// SIMATIC S7-200 project (STEP 7-Micro/WIN), CPU 224XP CN REL 02.01

SYMBOL_TABLE USER1
Pos_Real         VD100    // Posicion real en cuentas de encoder (REAL)
Setpoint         VD112    // Posicion objetivo de referencia en cuentas (REAL)
Accion_Control   VD116    // Accion de control calculada u (REAL)
K1               VD120    // Ganancia de posicion del controlador (97.7436) (REAL)
K2               VD124    // Ganancia de velocidad del controlador (25.8460) (REAL)
U_Abs            VD128    // Magnitud absoluta de la accion de control (REAL)
N                VD132    // Ganancia de precompensacion de la referencia (REAL)
Setpoint_In      VD136    // Referencia dinamica de posicion desde HMI (REAL)
Pos_Est          VD140    // Posicion estimada por el observador (REAL)
Vel_Est          VD144    // Velocidad estimada por el observador (REAL)
Error_Est        VD148    // Error de estimacion de la posicion ey (REAL)
L1               VD152    // Ganancia de observador para canal de posicion (0.1919) (REAL)
L2               VD156    // Ganancia de observador para canal de velocidad (0.6113) (REAL)
Phi12            VD160    // Matriz de transicion de estado elemento 12 (0.009814) (REAL)
Phi22            VD164    // Matriz de transicion de estado elemento 22 (0.963062) (REAL)
Gamma1           VD168    // Matriz de entrada elemento 1 (0.000008) (REAL)
Gamma2           VD172    // Matriz de entrada elemento 2 (0.001611) (REAL)
Pos_Est_Next     VD176    // Valor intermedio de posicion estimada siguiente (REAL)
Vel_Est_Next     VD180    // Valor intermedio de velocidad estimada siguiente (REAL)
Seta_Emergencia  I1.4     // Entrada de seguridad NC (1=OK
Variador_Run     Q0.0     // Mando Marcha/Paro del variador (1=Run
Variador_Dir     Q0.1     // Mando Direccion del variador (0=FWD
Salida_Analog    AQW0     // Consigna analoga de velocidad para el variador (0-32000)
Log_Pointer      VD400    // Puntero de escritura en la memoria de registro (DWORD)
Log_SampleCount  VW404    // Contador de muestras registradas de 0 a 200 (INT)
Log_DecimCount   VW406    // Contador de decimacion para muestreo de 50ms (INT)
Log_Active       V408.0   // Bandera de registro activo en ejecucion (BOOL)
Log_Trigger      V408.1   // Gatillo de inicio de registro manual (BOOL)
END_SYMBOL_TABLE

SYMBOL_TABLE S7-200 Symbols
Always_On        SM0.0    // 始终接通为 ON
First_Scan_On    SM0.1    // 仅第一个扫描周期中接通为 ON
Time_0_Intrvl    SMB34    // 定时中断 0 的时间间隔（从 1 至 255，以 1 毫秒为增量）。
HSC0_Ctrl        SMB37    // HSC0 设置与控制
HSC0_CV          SMD38    // HSC0 的新当前值
HSC0_PV          SMD42    // HSC0 的新预置值
END_SYMBOL_TABLE

ORGANIZATION_BLOCK MAIN:OB1
TITLE=
BEGIN
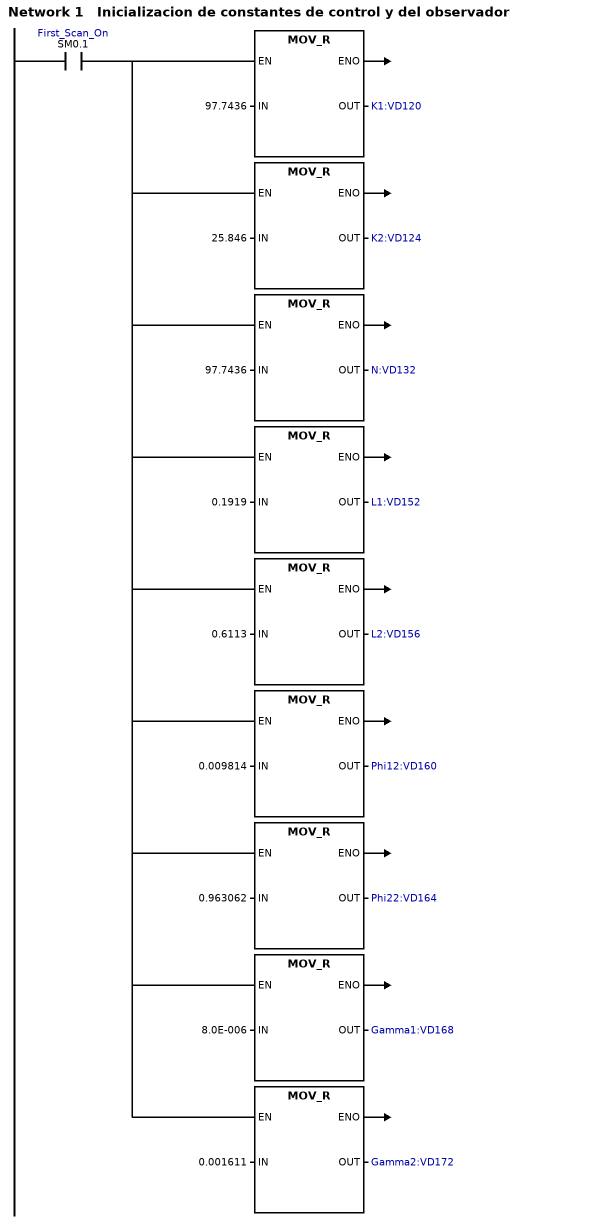
Network 1 //  Inicializacion de constantes de control y del observador
// K1
// K2
// N (Pre-compensacion)
// L1 (Ganancia de observador 1)
// L2 (Ganancia de observador 2)
// Phi12
// Phi22
// Gamma1
// Gamma2
LD     First_Scan_On:SM0.1
MOVR   97.7436, K1:VD120
MOVR   25.846, K2:VD124
MOVR   97.7436, N:VD132
MOVR   0.1919, L1:VD152
MOVR   0.6113, L2:VD156
MOVR   0.009814, Phi12:VD160
MOVR   0.963062, Phi22:VD164
MOVR   8.0E-006, Gamma1:VD168
MOVR   0.001611, Gamma2:VD172
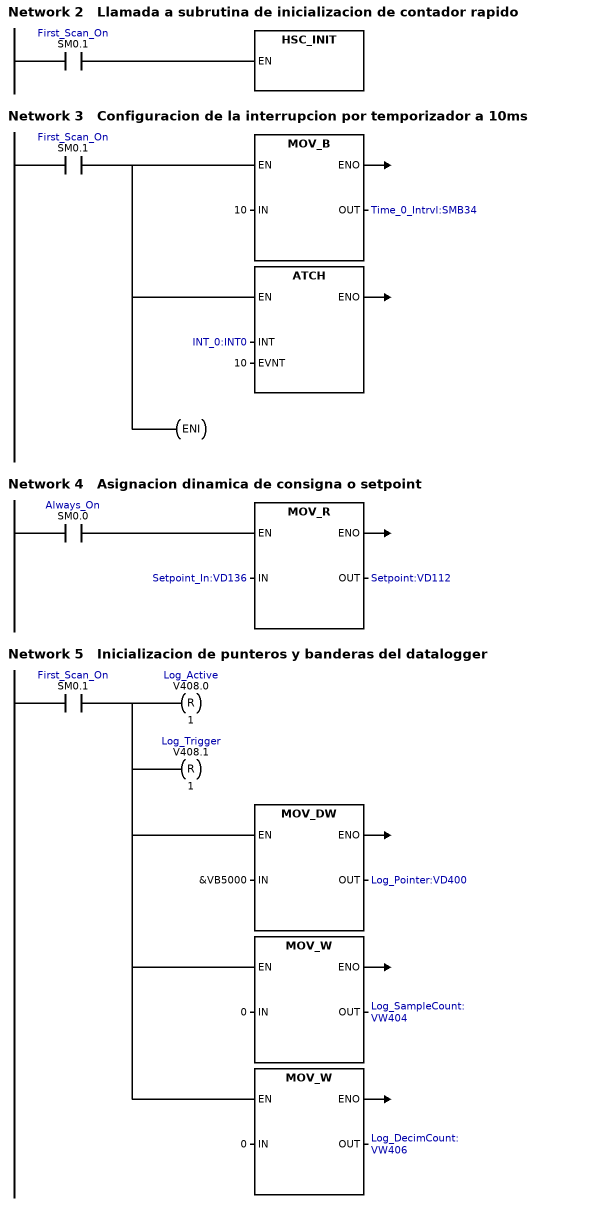
Network 2 //  Llamada a subrutina de inicializacion de contador rapido
// Llamada a SBR1 (HSC_INIT)
LD     First_Scan_On:SM0.1
CALL   HSC_INIT:SBR1
Network 3 //  Configuracion de la interrupcion por temporizador a 10ms
// Intervalo de interrupcion de 10ms
// Asociar INT0 al evento de temporizador 0
// Habilitar interrupciones globalmente
LD     First_Scan_On:SM0.1
MOVB   10, Time_0_Intrvl:SMB34
ATCH   INT_0:INT0, 10
ENI
Network 4 //  Asignacion dinamica de consigna o setpoint
// VD112 = Setpoint (Referencia)
LD     Always_On:SM0.0
MOVR   Setpoint_In:VD136, Setpoint:VD112
Network 5 //  Inicializacion de punteros y banderas del datalogger
// Desactivar bandera de datalogger activo
// Desactivar bandera de disparo (trigger)
// Direccion inicial del bufer en puntero
// Resetear contador de muestras
// Resetear contador de decimacion
LD     First_Scan_On:SM0.1
R      Log_Active:V408.0, 1
R      Log_Trigger:V408.1, 1
MOVD   &VB5000, Log_Pointer:VD400
MOVW   0, Log_SampleCount:VW404
MOVW   0, Log_DecimCount:VW406
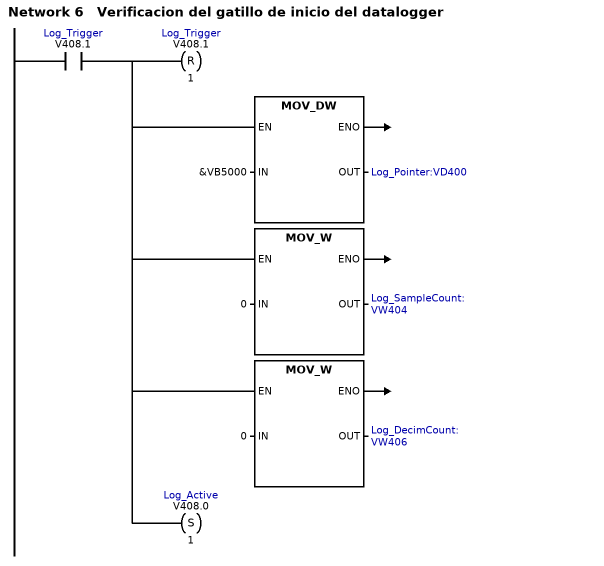
Network 6 //  Verificacion del gatillo de inicio del datalogger
// Si el usuario activa el gatillo
// Resetear bandera de gatillo
// Apuntar puntero al inicio VB5000
// Resetear contador de muestras
// Resetear contador de decimacion
// Activar bandera de datalogger activo
LD     Log_Trigger:V408.1
R      Log_Trigger:V408.1, 1
MOVD   &VB5000, Log_Pointer:VD400
MOVW   0, Log_SampleCount:VW404
MOVW   0, Log_DecimCount:VW406
S      Log_Active:V408.0, 1
END_ORGANIZATION_BLOCK

SUBROUTINE_BLOCK SBR_0:SBR0
TITLE=
BEGIN
Network 1
LD     Always_On:SM0.0
END_SUBROUTINE_BLOCK

SUBROUTINE_BLOCK HSC_INIT:SBR1
TITLE=
BEGIN
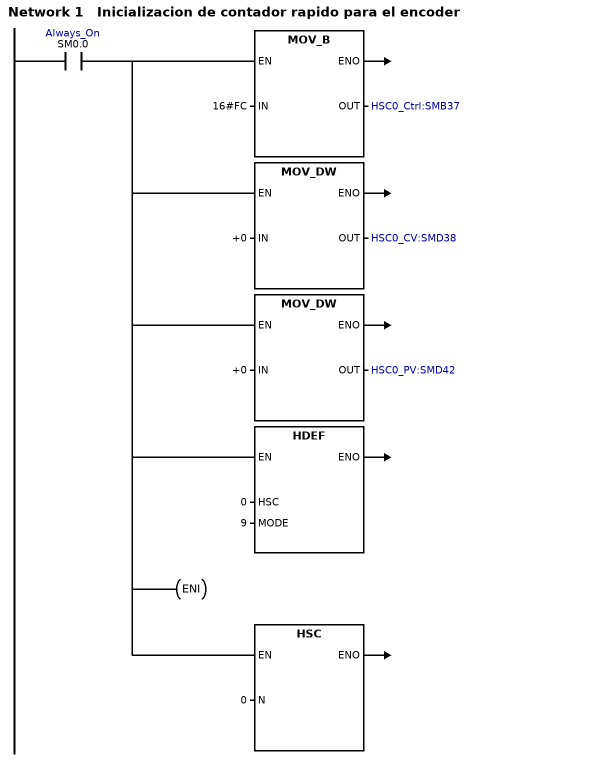
Network 1 //  Inicializacion de contador rapido para el encoder
// Configuracion de conteo: UP, 1X, habilitado
// Cargar valor actual (CV = 0)
// Cargar valor de preseleccion (PV = 0)
// Configurar HSC0 en Modo 9 (Fases A/B)
// Habilitar interrupciones
// Iniciar contador rapido HSC0
LD     Always_On:SM0.0
MOVB   16#FC, HSC0_Ctrl:SMB37
MOVD   +0, HSC0_CV:SMD38
MOVD   +0, HSC0_PV:SMD42
HDEF   0, 9
ENI
HSC    0
END_SUBROUTINE_BLOCK

INTERRUPT_BLOCK INT_0:INT0
TITLE=
BEGIN
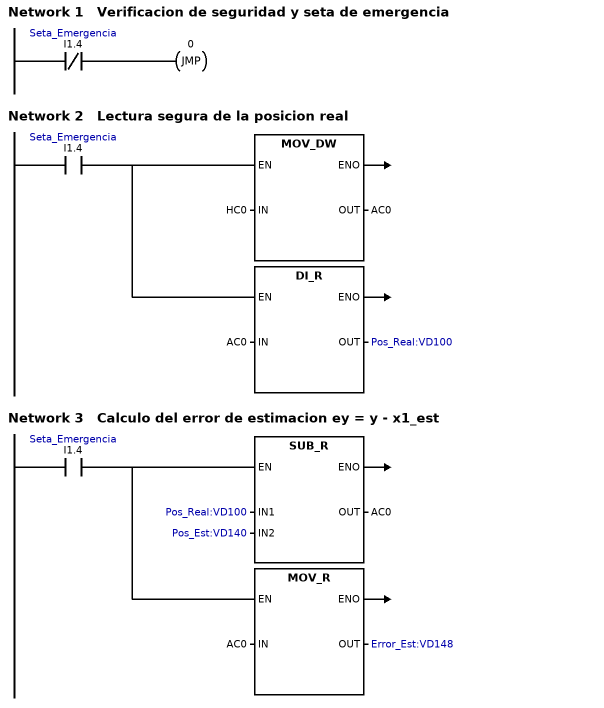
Network 1 //  Verificacion de seguridad y seta de emergencia
// Si la seta de emergencia se activa (NC abierto)
// Saltar a la etiqueta de parada segura
LDN    Seta_Emergencia:I1.4
JMP    0
Network 2 //  Lectura segura de la posicion real
// Mover lectura de HC0 a AC0
// Convertir entero de AC0 a REAL en VD100 (y)
LD     Seta_Emergencia:I1.4
MOVD   HC0, AC0
DTR    AC0, Pos_Real:VD100
Network 3 //  Calculo del error de estimacion ey = y - x1_est
// AC0 = y
// AC0 = y - x1_est
// VD148 = ey
LD     Seta_Emergencia:I1.4
MOVR   Pos_Real:VD100, AC0
-R     Pos_Est:VD140, AC0
MOVR   AC0, Error_Est:VD148
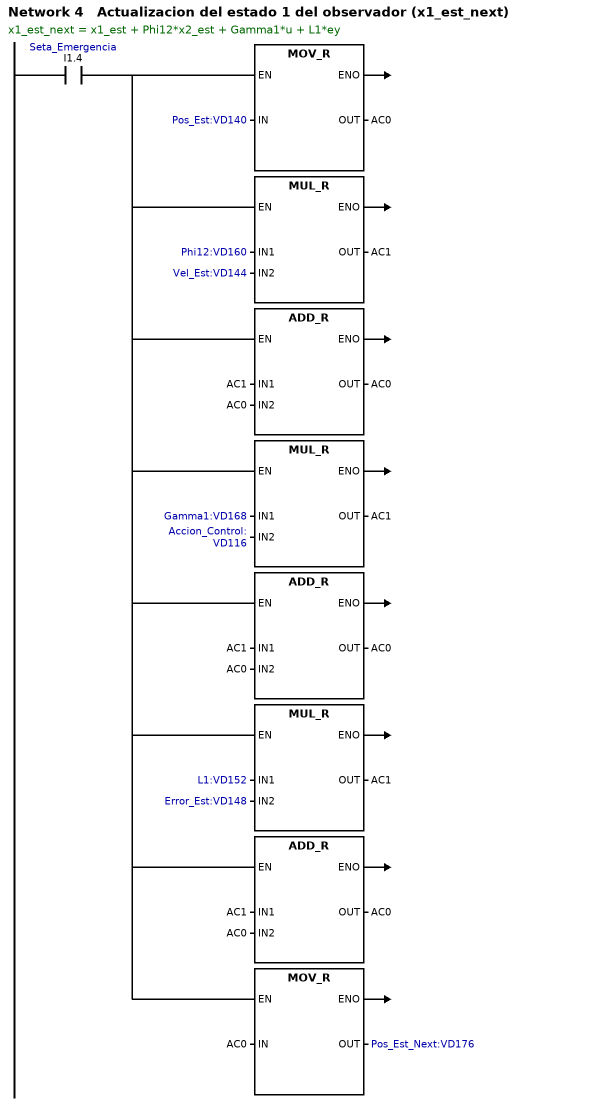
Network 4 //  Actualizacion del estado 1 del observador (x1_est_next)
//  x1_est_next = x1_est + Phi12*x2_est + Gamma1*u + L1*ey
// AC0 = x1_est
// AC1 = Phi12
// AC1 = Phi12 * x2_est
// AC0 = x1_est + Phi12*x2_est
// AC1 = Gamma1
// AC1 = Gamma1 * u
// AC1 = L1
// AC1 = L1 * ey
// VD176 = x1_est_next (temporal)
LD     Seta_Emergencia:I1.4
MOVR   Pos_Est:VD140, AC0
MOVR   Phi12:VD160, AC1
*R     Vel_Est:VD144, AC1
+R     AC1, AC0
MOVR   Gamma1:VD168, AC1
*R     Accion_Control:VD116, AC1
+R     AC1, AC0
MOVR   L1:VD152, AC1
*R     Error_Est:VD148, AC1
+R     AC1, AC0
MOVR   AC0, Pos_Est_Next:VD176
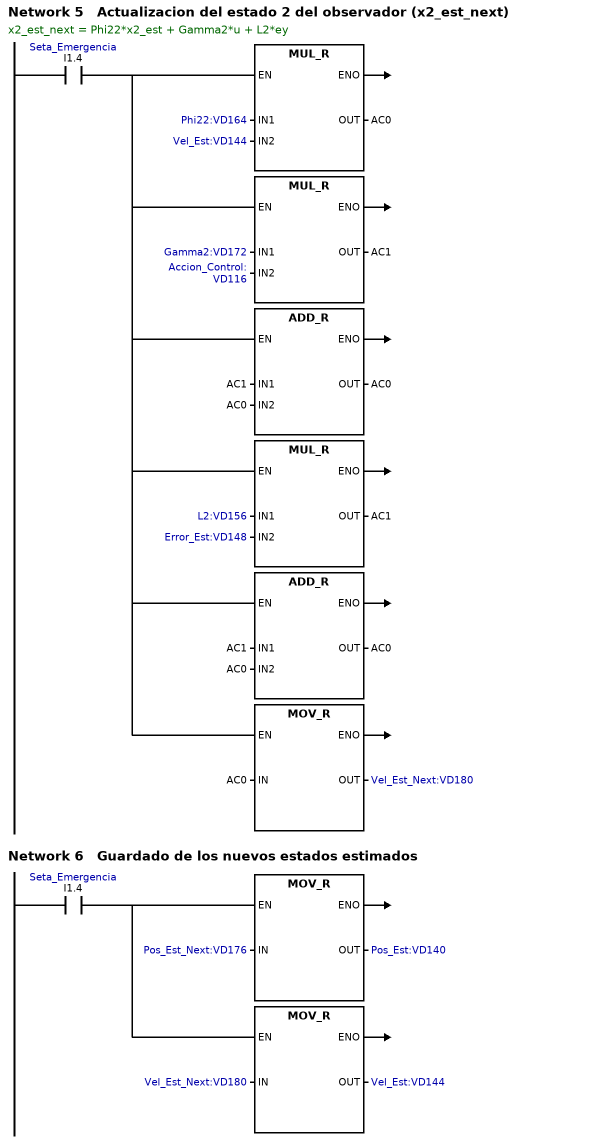
Network 5 //  Actualizacion del estado 2 del observador (x2_est_next)
//  x2_est_next = Phi22*x2_est + Gamma2*u + L2*ey
// AC0 = Phi22
// AC0 = Phi22 * x2_est
// AC1 = Gamma2
// AC1 = Gamma2 * u
// AC1 = L2
// AC1 = L2 * ey
// VD180 = x2_est_next (temporal)
LD     Seta_Emergencia:I1.4
MOVR   Phi22:VD164, AC0
*R     Vel_Est:VD144, AC0
MOVR   Gamma2:VD172, AC1
*R     Accion_Control:VD116, AC1
+R     AC1, AC0
MOVR   L2:VD156, AC1
*R     Error_Est:VD148, AC1
+R     AC1, AC0
MOVR   AC0, Vel_Est_Next:VD180
Network 6 //  Guardado de los nuevos estados estimados
// Actualizar x1_est
// Actualizar x2_est
LD     Seta_Emergencia:I1.4
MOVR   Pos_Est_Next:VD176, Pos_Est:VD140
MOVR   Vel_Est_Next:VD180, Vel_Est:VD144
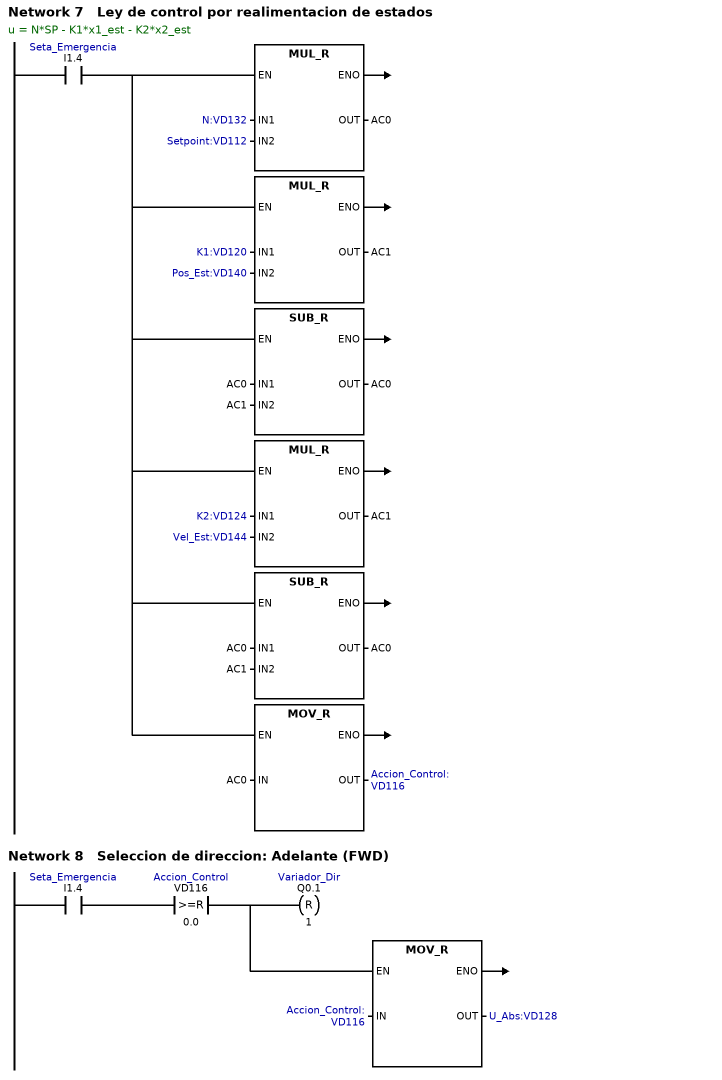
Network 7 //  Ley de control por realimentacion de estados
//  u = N*SP - K1*x1_est - K2*x2_est
// AC0 = N
// AC0 = N * SP
// AC1 = K1
// AC1 = K1 * x1_est
// AC0 = N*SP - K1*x1_est
// AC1 = K2
// AC1 = K2 * x2_est
// AC0 = u final
// VD116 = Accion de Control (u)
LD     Seta_Emergencia:I1.4
MOVR   N:VD132, AC0
*R     Setpoint:VD112, AC0
MOVR   K1:VD120, AC1
*R     Pos_Est:VD140, AC1
-R     AC1, AC0
MOVR   K2:VD124, AC1
*R     Vel_Est:VD144, AC1
-R     AC1, AC0
MOVR   AC0, Accion_Control:VD116
Network 8 //  Seleccion de direccion: Adelante (FWD)
// Si u >= 0
// Desactivar sentido inverso (FWD)
// Copiar magnitud a VD128
LD     Seta_Emergencia:I1.4
AR>=   Accion_Control:VD116, 0.0
R      Variador_Dir:Q0.1, 1
MOVR   Accion_Control:VD116, U_Abs:VD128
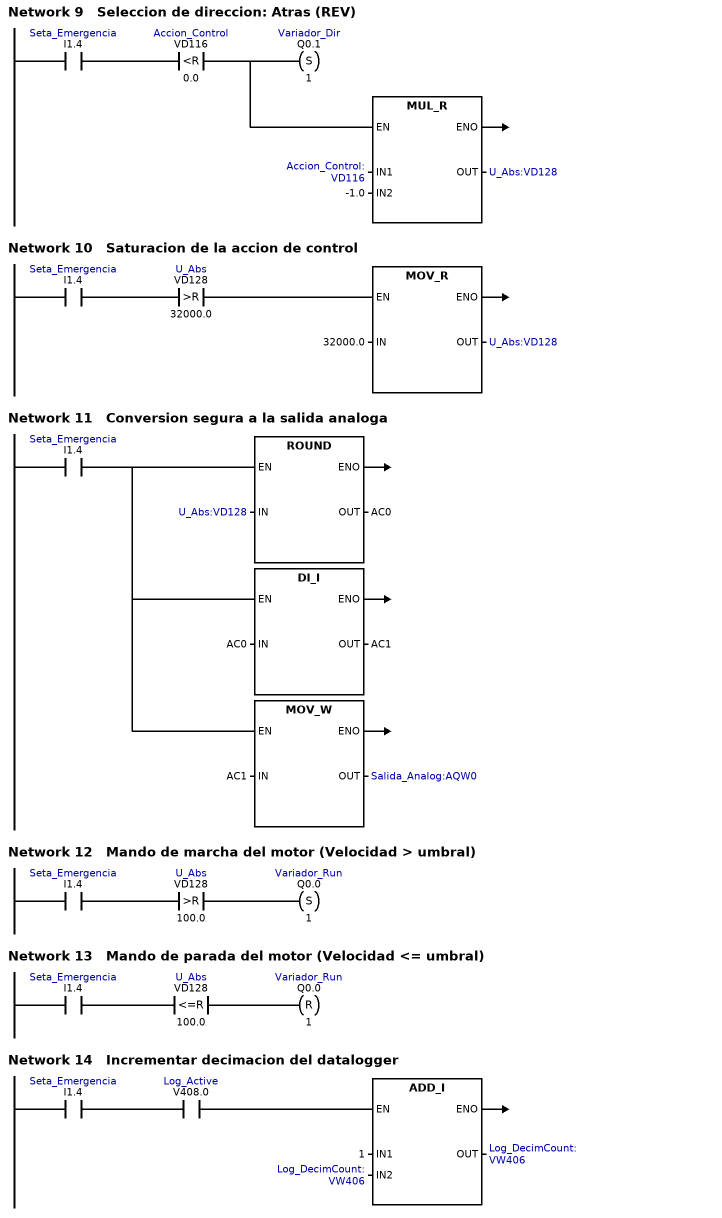
Network 9 //  Seleccion de direccion: Atras (REV)
// Si u < 0
// Activar sentido inverso (REV)
// Copiar magnitud absoluta |u| a VD128
LD     Seta_Emergencia:I1.4
AR<    Accion_Control:VD116, 0.0
S      Variador_Dir:Q0.1, 1
MOVR   Accion_Control:VD116, U_Abs:VD128
*R     -1.0, U_Abs:VD128
Network 10 //  Saturacion de la accion de control
// Si la magnitud supera los 10V
// Limitar consigna a 32000
LD     Seta_Emergencia:I1.4
AR>    U_Abs:VD128, 32000.0
MOVR   32000.0, U_Abs:VD128
Network 11 //  Conversion segura a la salida analoga
// Redondear REAL a DINT en AC0
// Convertir DINT a INT en AC1
// Escribir Word en la salida analoga
LD     Seta_Emergencia:I1.4
ROUND  U_Abs:VD128, AC0
DTI    AC0, AC1
MOVW   AC1, Salida_Analog:AQW0
Network 12 //  Mando de marcha del motor (Velocidad > umbral)
// Si supera la zona muerta
// Arrancar motor (RUN)
LD     Seta_Emergencia:I1.4
AR>    U_Abs:VD128, 100.0
S      Variador_Run:Q0.0, 1
Network 13 //  Mando de parada del motor (Velocidad <= umbral)
// Si cae dentro de la zona muerta
// Parar motor (STOP)
LD     Seta_Emergencia:I1.4
AR<=   U_Abs:VD128, 100.0
R      Variador_Run:Q0.0, 1
Network 14 //  Incrementar decimacion del datalogger
// Si el registro esta activo
// Incrementar decimacion
LD     Seta_Emergencia:I1.4
A      Log_Active:V408.0
+I     1, Log_DecimCount:VW406
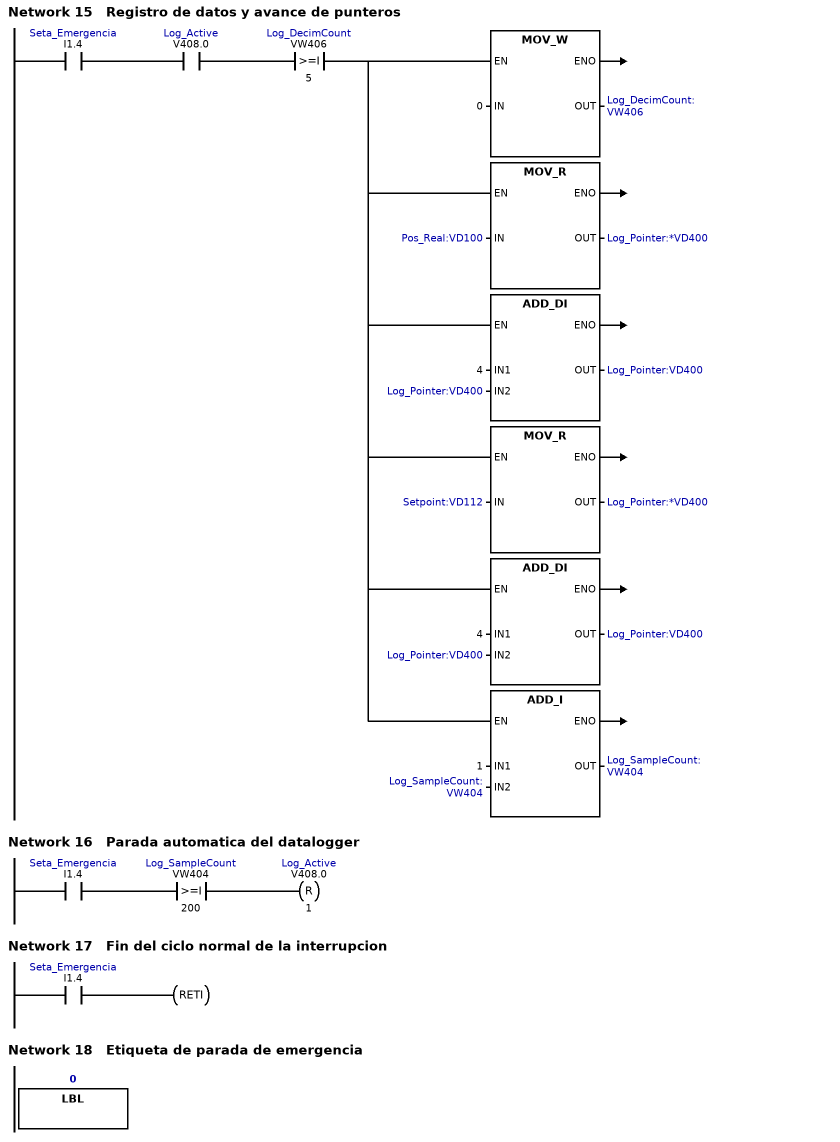
Network 15 //  Registro de datos y avance de punteros
// Si han pasado 50ms
// Resetear decimacion
// Guardar posicion real
// Avanzar puntero a setpoint
// Guardar setpoint
// Avanzar puntero a posicion siguiente
// Incrementar contador de muestras
LD     Seta_Emergencia:I1.4
A      Log_Active:V408.0
AW>=   Log_DecimCount:VW406, 5
MOVW   0, Log_DecimCount:VW406
MOVR   Pos_Real:VD100, *Log_Pointer:VD400
+D     4, Log_Pointer:VD400
MOVR   Setpoint:VD112, *Log_Pointer:VD400
+D     4, Log_Pointer:VD400
+I     1, Log_SampleCount:VW404
Network 16 //  Parada automatica del datalogger
// Si se alcanza el limite de 200 muestras
// Detener adquisicion
LD     Seta_Emergencia:I1.4
AW>=   Log_SampleCount:VW404, 200
R      Log_Active:V408.0, 1
Network 17 //  Fin del ciclo normal de la interrupcion
// Retorno de interrupcion
LD     Seta_Emergencia:I1.4
CRETI
Network 18 //  Etiqueta de parada de emergencia
LBL    0
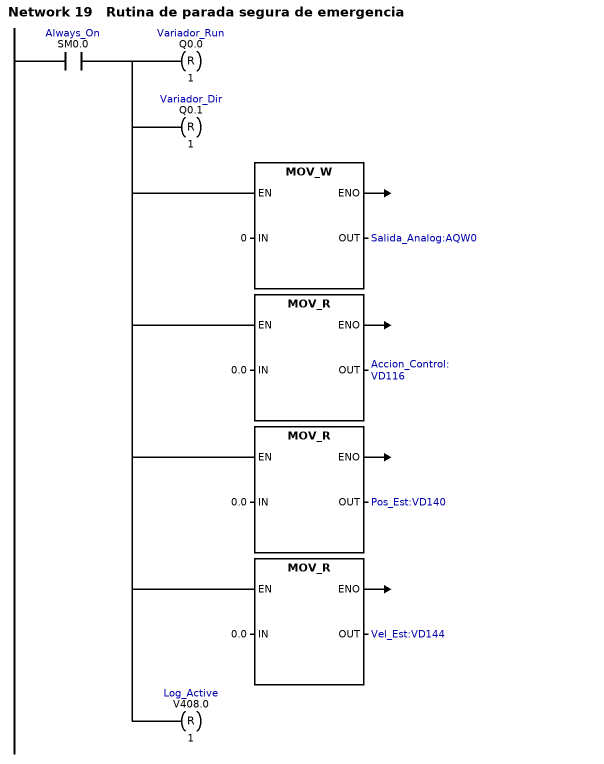
Network 19 //  Rutina de parada segura de emergencia
// Apagar motor inmediatamente
// Desactivar sentido de giro
// Escribir cero en salida analoga
// Resetear accion de control
// Resetear posicion estimada
// Resetear velocidad estimada
// Apagar datalogger
LD     Always_On:SM0.0
R      Variador_Run:Q0.0, 1
R      Variador_Dir:Q0.1, 1
MOVW   0, Salida_Analog:AQW0
MOVR   0.0, Accion_Control:VD116
MOVR   0.0, Pos_Est:VD140
MOVR   0.0, Vel_Est:VD144
R      Log_Active:V408.0, 1
END_INTERRUPT_BLOCK
